Fanuc TP program (LS listing): SplitTest.LS

/PROG  SplitTest
/ATTR
OWNER		= MNEDITOR;
COMMENT		= "RoboDK sequence";
PROG_SIZE	= 0;
CREATE		= DATE 31-12-14  TIME 12:00:00;
MODIFIED	= DATE 31-12-14  TIME 12:00:00;
FILE_NAME	= SplitTest;
VERSION		= 0;
LINE_COUNT	= 15;
MEMORY_SIZE	= 0;
PROTECT		= READ_WRITE;
TCD:  STACK_SIZE	= 0,
      TASK_PRIORITY	= 50,
      TIME_SLICE	= 0,
      BUSY_LAMP_OFF	= 0,
      ABORT_REQUEST	= 0,
      PAUSE_REQUEST	= 0;
DEFAULT_GROUP	= 1,*,*,*,*,*,*;
CONTROL_CODE	= 00000000 00000000;
/MN
   1:  ! Program generated by VerticalBot Studio for Fanuc LR Mate 200 ;
   2:  ! iD on 25/10/2026 12:00:00 ;
   3:  ! Using nominal kinematics. ;
   4:  UFRAME_NUM=2 ;
   5:  ! UF2:100.0,-50.0,20.0,0.0,0.0,30.0 ;
   6:  UTOOL_NUM=1 ;
   7:  ! UT1:10.0,0.0,120.0,0.0,15.0,0.0 ;
   8:J P[1] 4% FINE ;
   9:L P[2] 200mm/sec FINE ;
  10:L P[3] 200mm/sec FINE ;
  11:L P[4] 200mm/sec FINE ;
  12:L P[5] 200mm/sec FINE ;
  13:L P[6] 200mm/sec FINE ;
  14:L P[7] 200mm/sec FINE ;
  15:L P[8] 200mm/sec FINE ;
/POS
P[1]{
   GP1:
    UF : 2, UT : 1,
	J1=    -20.000 deg,	J2=    10.000 deg,	J3=    -20.000 deg,
	J4=    30.000 deg,	J5=    -40.000 deg,	J6=    50.000 deg
};
P[2]{
   GP1:
    UF : 2, UT : 1,        CONFIG : 'F U T, 0, 0, 0',
	X =   332.153  mm,	Y =  -359.974  mm,	Z =   826.762  mm,
	W =   -51.647 deg,	P =     9.441 deg,	R =  -168.258 deg
};
P[3]{
   GP1:
    UF : 2, UT : 1,        CONFIG : 'F U T, 0, 0, 0',
	X =   286.258  mm,	Y =  -372.547  mm,	Z =   823.386  mm,
	W =   -52.463 deg,	P =     8.848 deg,	R =  -172.388 deg
};
P[4]{
   GP1:
    UF : 2, UT : 1,        CONFIG : 'F U T, 0, 0, 0',
	X =   332.153  mm,	Y =  -359.974  mm,	Z =   826.762  mm,
	W =   -51.647 deg,	P =     9.441 deg,	R =  -168.258 deg
};
P[5]{
   GP1:
    UF : 2, UT : 1,        CONFIG : 'F U T, 0, 0, 0',
	X =   286.258  mm,	Y =  -372.547  mm,	Z =   823.386  mm,
	W =   -52.463 deg,	P =     8.848 deg,	R =  -172.388 deg
};
P[6]{
   GP1:
    UF : 2, UT : 1,        CONFIG : 'F U T, 0, 0, 0',
	X =   332.153  mm,	Y =  -359.974  mm,	Z =   826.762  mm,
	W =   -51.647 deg,	P =     9.441 deg,	R =  -168.258 deg
};
P[7]{
   GP1:
    UF : 2, UT : 1,        CONFIG : 'F U T, 0, 0, 0',
	X =   286.258  mm,	Y =  -372.547  mm,	Z =   823.386  mm,
	W =   -52.463 deg,	P =     8.848 deg,	R =  -172.388 deg
};
P[8]{
   GP1:
    UF : 2, UT : 1,        CONFIG : 'F U T, 0, 0, 0',
	X =   332.153  mm,	Y =  -359.974  mm,	Z =   826.762  mm,
	W =   -51.647 deg,	P =     9.441 deg,	R =  -168.258 deg
};
/END
